(* IEC 61131-3 sources: volt/packages/volt-lsp-iec/test-corpus/lenze-mid/Device/Plc Logic/Application/Library Manager/CAA MemBlockMan, 94 files *)

(* ---- BCP.dut ---- *)
TYPE BCP :
STRUCT
	PPOOL : POINTER TO PCB;
END_STRUCT
END_TYPE

(* ---- ERROR.dut ---- *)
TYPE ERROR :
(
	NO_ERROR := 0,
	FIRST_ERROR := 30100,
	UNKNOWN_EVENT := 30102,
	NOMORE_MEMORY := 30103,
	WRONG_PRIO := 30104,
	EMPTY_LIST := 30105,
	NO_EXIST_PRIO := 30106,
	PRIO_EXIST := 30107,
	PRIOS_EXCEED := 30108,
	ALIGNMENT_ERROR := 30109,
	BLOCKSIZE_TO_SMALL := 30110,
	EMPTY_POOL := 30111,
	EMPTY_EXCHANGE := 30112,
	TIMEOUT := 30113,
	WRONG_TIMEOUT := 30114,
	REF_OVERFLOW := 30115,
	WRONG_KEY := 30116,
	HANDLE_INVALID := 30117,
	REF_NOT_ZERO := 30118,
	WRONG_NUM_OF_MSG := 30119,
	BUFFER_TO_BIG := 30120,
	WRONG_OP := 30121,
	GEN_ERROR := 30149,
	FIRST_MF := 30150,
	LAST_ERROR := 30199
);
END_TYPE

(* ---- PCB.dut ---- *)
TYPE PCB :
STRUCT
	XWDUMMYA : __XWORD;
	SZBLOCK : CAA.SIZE;
	XWDUMMYB : __XWORD;
	XWDUMMYC : __XWORD;
	CTBLKLEFT : CAA.COUNT;
	CTBLKCAP : CAA.COUNT;
END_STRUCT
END_TYPE

(* ---- RSHANDLING.gvl ---- *)
VAR_GLOBAL
	G_XCHGCLASS : XChgClass;
	G_FLATCLASS : FlatClass;
	G_MSGCLASS : MsgClass;
	G_REFCLASS : MsgClass;
	G_POOLCLASS : PoolClass;
	G_BLKCLASS : BlkClass;
	G_RLSTCLASS : RLstClass;
END_VAR

(* ---- VERSIONCONSTANTS.gvl ---- *)
VAR_GLOBAL
	GC_BYVERSION : BYTE := 1;
	GC_VERSION_1 : BYTE := 0;
END_VAR

(* ---- _BLOCKGETDATA.pou ---- *)
FUNCTION _BLOCKGETDATA : CAA.PVOID
VAR_INPUT
	HBLOCK : CAA.HANDLE;
	PEERROR : POINTER TO ERROR;
END_VAR
END_FUNCTION

(* ---- _BLOCKGETPOOL.pou ---- *)
FUNCTION _BLOCKGETPOOL : CAA.HANDLE
VAR_INPUT
	HBLOCK : CAA.HANDLE;
	PEERROR : POINTER TO ERROR;
END_VAR
END_FUNCTION

(* ---- _FLATCREATEH.pou ---- *)
FUNCTION _FLATCREATEH : CAA.HANDLE
VAR_INPUT
	IDMINKEY : CAA.IDENT;
	IDMAXKEY : CAA.IDENT;
	CTNUMKEYS : CAA.COUNT;
	EENABLE : CB.EVENT;
	EDISABLE : CB.EVENT;
	EUPDATE : CB.EVENT;
	EREAD : CB.EVENT;
	PEERROR : POINTER TO ERROR;
END_VAR
END_FUNCTION

(* ---- _FLATCREATEP.pou ---- *)
FUNCTION _FLATCREATEP : CAA.HANDLE
VAR_INPUT
	IDMINKEY : CAA.IDENT;
	IDMAXKEY : CAA.IDENT;
	CTNUMKEY : CAA.COUNT;
	SZMEMSIZE : CAA.SIZE;
	PMEMORY : CAA.PVOID;
	EENABLE : CB.EVENT;
	EDISABLE : CB.EVENT;
	EUPDATE : CB.EVENT;
	EREAD : CB.EVENT;
	PEERROR : POINTER TO ERROR;
END_VAR
END_FUNCTION

(* ---- _FLATDELETE.pou ---- *)
FUNCTION _FLATDELETE : ERROR
VAR_INPUT
	HFLAT : CAA.HANDLE;
END_VAR
END_FUNCTION

(* ---- _FLATDISABLE.pou ---- *)
FUNCTION _FLATDISABLE : CAA.HANDLE
VAR_INPUT
	HFLAT : CAA.HANDLE;
	IDKEY : CAA.IDENT;
	PEERROR : POINTER TO ERROR;
END_VAR
END_FUNCTION

(* ---- _FLATENABLE.pou ---- *)
FUNCTION _FLATENABLE : ERROR
VAR_INPUT
	HFLAT : CAA.HANDLE;
	IDKEY : CAA.IDENT;
END_VAR
END_FUNCTION

(* ---- _FLATGETSIZE.pou ---- *)
FUNCTION _FLATGETSIZE : CAA.SIZE
VAR_INPUT
	CTNUMKEYS : CAA.COUNT;
END_VAR
END_FUNCTION

(* ---- _FLATREAD.pou ---- *)
FUNCTION _FLATREAD : CAA.HANDLE
VAR_INPUT
	HFLAT : CAA.HANDLE;
	IDKEY : CAA.IDENT;
	PEERROR : POINTER TO ERROR;
END_VAR
END_FUNCTION

(* ---- _FLATTEST.pou ---- *)
FUNCTION _FLATTEST : BOOL
VAR_INPUT
	HFLAT : CAA.HANDLE;
	IDKEY : CAA.IDENT;
	PEERROR : POINTER TO ERROR;
END_VAR
END_FUNCTION

(* ---- _FLATUPDATE.pou ---- *)
FUNCTION _FLATUPDATE : CAA.HANDLE
VAR_INPUT
	HFLAT : CAA.HANDLE;
	IDKEY : CAA.IDENT;
	HMSG : CAA.HANDLE;
	PEERROR : POINTER TO ERROR;
END_VAR
END_FUNCTION

(* ---- _MSGADDREF.pou ---- *)
FUNCTION _MSGADDREF : ERROR
VAR_INPUT
	HMSG : CAA.HANDLE;
END_VAR
END_FUNCTION

(* ---- _MSGCLONE.pou ---- *)
FUNCTION _MSGCLONE : CAA.HANDLE
VAR_INPUT
	HMSG : CAA.HANDLE;
	PEERROR : POINTER TO ERROR;
END_VAR
END_FUNCTION

(* ---- _MSGGETDATA.pou ---- *)
FUNCTION _MSGGETDATA : CAA.PVOID
VAR_INPUT
	HMSG : CAA.HANDLE;
	PEERROR : POINTER TO ERROR;
END_VAR
END_FUNCTION

(* ---- _MSGRECEIVE.pou ---- *)
FUNCTION _MSGRECEIVE : CAA.HANDLE
VAR_INPUT
	HXCHG : CAA.HANDLE;
	PCTMSGLEFT : POINTER TO CAA.COUNT;
	PEERROR : POINTER TO ERROR;
END_VAR
END_FUNCTION

(* ---- _MSGRELEASE.pou ---- *)
FUNCTION _MSGRELEASE : ERROR
VAR_INPUT
	HMSG : CAA.HANDLE;
END_VAR
END_FUNCTION

(* ---- _MSGRELEASEEX.pou ---- *)
FUNCTION _MSGRELEASEEX : ERROR
VAR_INPUT
	HMSG : CAA.HANDLE;
	HXCHG : CAA.HANDLE;
END_VAR
END_FUNCTION

(* ---- _MSGSEND.pou ---- *)
FUNCTION _MSGSEND : ERROR
VAR_INPUT
	HMSG : CAA.HANDLE;
	USIPRIO : USINT;
	HXCHG : CAA.HANDLE;
END_VAR
END_FUNCTION

(* ---- _POOLCREATEH.pou ---- *)
FUNCTION _POOLCREATEH : CAA.HANDLE
VAR_INPUT
	CTNUMBLOCKS : CAA.COUNT;
	SZBLOCKSIZE : CAA.SIZE;
	EEMPTY : CB.EVENT;
	PEERROR : POINTER TO ERROR;
END_VAR
END_FUNCTION

(* ---- _POOLCREATEP.pou ---- *)
FUNCTION _POOLCREATEP : CAA.HANDLE
VAR_INPUT
	SZBLOCKSIZE : CAA.SIZE;
	SZMEMSIZE : CAA.SIZE;
	PMEMORY : CAA.PVOID;
	EEMPTY : CB.EVENT;
	PEERROR : POINTER TO ERROR;
END_VAR
END_FUNCTION

(* ---- _POOLDELETE.pou ---- *)
FUNCTION _POOLDELETE : ERROR
VAR_INPUT
	HPOOL : CAA.HANDLE;
END_VAR
END_FUNCTION

(* ---- _POOLEXTENDH.pou ---- *)
FUNCTION _POOLEXTENDH : ERROR
VAR_INPUT
	HPOOL : CAA.HANDLE;
	CTNUMBLOCKS : CAA.COUNT;
END_VAR
END_FUNCTION

(* ---- _POOLGETBLOCK.pou ---- *)
FUNCTION _POOLGETBLOCK : CAA.HANDLE
VAR_INPUT
	HPOOL : CAA.HANDLE;
	PEERROR : POINTER TO ERROR;
END_VAR
END_FUNCTION

(* ---- _POOLGETBLOCKSIZE.pou ---- *)
FUNCTION _POOLGETBLOCKSIZE : CAA.SIZE
VAR_INPUT
	HPOOL : CAA.HANDLE;
	PEERROR : POINTER TO ERROR;
END_VAR
END_FUNCTION

(* ---- _POOLGETCURCAPACITY.pou ---- *)
FUNCTION _POOLGETCURCAPACITY : CAA.COUNT
VAR_INPUT
	HPOOL : CAA.HANDLE;
	PEERROR : POINTER TO ERROR;
END_VAR
END_FUNCTION

(* ---- _POOLGETNUMBLOCKSLEFT.pou ---- *)
FUNCTION _POOLGETNUMBLOCKSLEFT : CAA.COUNT
VAR_INPUT
	HPOOL : CAA.HANDLE;
	PEERROR : POINTER TO ERROR;
END_VAR
END_FUNCTION

(* ---- _POOLGETSIZE.pou ---- *)
FUNCTION _POOLGETSIZE : CAA.SIZE
VAR_INPUT
	CTNUMBLOCK : CAA.COUNT;
	SZBLOCKSIZE : CAA.SIZE;
END_VAR
END_FUNCTION

(* ---- _POOLPUTBLOCK.pou ---- *)
FUNCTION _POOLPUTBLOCK : ERROR
VAR_INPUT
	HBLOCK : CAA.HANDLE;
END_VAR
END_FUNCTION

(* ---- _RLSTADDPRIO.pou ---- *)
FUNCTION _RLSTADDPRIO : ERROR
VAR_INPUT
	HRLST : CAA.HANDLE;
	USIPRIO : USINT;
END_VAR
END_FUNCTION

(* ---- _RLSTCHECKPRIO.pou ---- *)
FUNCTION _RLSTCHECKPRIO : BOOL
VAR_INPUT
	HRLST : CAA.HANDLE;
	USIPRIO : USINT;
	PEERROR : POINTER TO ERROR;
END_VAR
END_FUNCTION

(* ---- _RLSTCREATEH.pou ---- *)
FUNCTION _RLSTCREATEH : CAA.HANDLE
VAR_INPUT
	PEERROR : POINTER TO ERROR;
END_VAR
END_FUNCTION

(* ---- _RLSTCREATEP.pou ---- *)
FUNCTION _RLSTCREATEP : CAA.HANDLE
VAR_INPUT
	SZMEMORY : CAA.SIZE;
	PMEMORY : CAA.PVOID;
	PEERROR : POINTER TO ERROR;
END_VAR
END_FUNCTION

(* ---- _RLSTDELETE.pou ---- *)
FUNCTION _RLSTDELETE : ERROR
VAR_INPUT
	HRLST : CAA.HANDLE;
END_VAR
END_FUNCTION

(* ---- _RLSTGETHIGHESTPRIO.pou ---- *)
FUNCTION _RLSTGETHIGHESTPRIO : USINT
VAR_INPUT
	HRLST : CAA.HANDLE;
	PEERROR : POINTER TO ERROR;
END_VAR
END_FUNCTION

(* ---- _RLSTGETSIZE.pou ---- *)
FUNCTION _RLSTGETSIZE : CAA.SIZE
VAR_INPUT
	XDUMMY : BOOL;
END_VAR
END_FUNCTION

(* ---- _RLSTREMOVEPRIO.pou ---- *)
FUNCTION _RLSTREMOVEPRIO : ERROR
VAR_INPUT
	HRLST : CAA.HANDLE;
	USIPRIO : USINT;
END_VAR
END_FUNCTION

(* ---- _XCHGCREATEH.pou ---- *)
FUNCTION _XCHGCREATEH : CAA.HANDLE
VAR_INPUT
	CTNUMMSG : CAA.COUNT;
	SZBLOCKSIZE : CAA.SIZE;
	CTNUMPRIOS : CAA.COUNT;
	ESENDMSG : CB.EVENT;
	ERECEIVEMSG : CB.EVENT;
	EXCHGEMPTY : CB.EVENT;
	PEERROR : POINTER TO ERROR;
END_VAR
END_FUNCTION

(* ---- _XCHGCREATEP.pou ---- *)
FUNCTION _XCHGCREATEP : CAA.HANDLE
VAR_INPUT
	SZBLOCKSIZE : CAA.SIZE;
	CTNUMPRIOS : CAA.COUNT;
	SZMEMSIZE : CAA.SIZE;
	PMEMORY : CAA.PVOID;
	ESENDMSG : CB.EVENT;
	ERECEIVEMSG : CB.EVENT;
	EXCHGEMPTY : CB.EVENT;
	PEERROR : POINTER TO ERROR;
END_VAR
END_FUNCTION

(* ---- _XCHGDELETE.pou ---- *)
FUNCTION _XCHGDELETE : ERROR
VAR_INPUT
	HXCHG : CAA.HANDLE;
END_VAR
END_FUNCTION

(* ---- _XCHGEXTENDH.pou ---- *)
FUNCTION _XCHGEXTENDH : ERROR
VAR_INPUT
	HXCHG : CAA.HANDLE;
	CTNUMMSG : CAA.COUNT;
END_VAR
END_FUNCTION

(* ---- _XCHGGETSIZE.pou ---- *)
FUNCTION _XCHGGETSIZE : CAA.SIZE
VAR_INPUT
	CTNUMMSG : CAA.COUNT;
	SZBLOCKSIZE : CAA.SIZE;
	CTNUMPRIOS : CAA.COUNT;
END_VAR
END_FUNCTION

(* ---- _XCHGISEMPTY.pou ---- *)
FUNCTION _XCHGISEMPTY : BOOL
VAR_INPUT
	HXCHG : CAA.HANDLE;
	PEERROR : POINTER TO ERROR;
END_VAR
END_FUNCTION

(* ---- _XCHGMSGLEFT.pou ---- *)
FUNCTION _XCHGMSGLEFT : CAA.COUNT
VAR_INPUT
	HXCHG : CAA.HANDLE;
	PEERROR : POINTER TO ERROR;
END_VAR
END_FUNCTION

(* ---- BLOCKGETDATA.pou ---- *)
FUNCTION BLOCKGETDATA : CAA.PVOID
VAR_INPUT
	HBLOCK : CAA.HANDLE;
	PEERROR : POINTER TO ERROR;
END_VAR
END_FUNCTION

(* ---- FLATCREATEH.pou ---- *)
FUNCTION FLATCREATEH : CAA.HANDLE
VAR_INPUT
	IDMINKEY : CAA.IDENT;
	IDMAXKEY : CAA.IDENT;
	CTNUMKEYS : CAA.COUNT;
	EENABLE : CB.EVENT;
	EDISABLE : CB.EVENT;
	EUPDATE : CB.EVENT;
	EREAD : CB.EVENT;
	PEERROR : POINTER TO ERROR;
END_VAR
END_FUNCTION

(* ---- FLATCREATEP.pou ---- *)
FUNCTION FLATCREATEP : CAA.HANDLE
VAR_INPUT
	IDMINKEY : CAA.IDENT;
	IDMAXKEY : CAA.IDENT;
	CTNUMKEY : CAA.COUNT;
	SZMEMSIZE : CAA.SIZE;
	PMEMORY : CAA.PVOID;
	EENABLE : CB.EVENT;
	EDISABLE : CB.EVENT;
	EUPDATE : CB.EVENT;
	EREAD : CB.EVENT;
	PEERROR : POINTER TO ERROR;
END_VAR
END_FUNCTION

(* ---- FLATDELETE.pou ---- *)
FUNCTION FLATDELETE : ERROR
VAR_INPUT
	HFLAT : CAA.HANDLE;
END_VAR
END_FUNCTION

(* ---- FLATDISABLE.pou ---- *)
FUNCTION FLATDISABLE : CAA.HANDLE
VAR_INPUT
	HFLAT : CAA.HANDLE;
	IDKEY : CAA.IDENT;
	PEERROR : POINTER TO ERROR;
END_VAR
END_FUNCTION

(* ---- FLATENABLE.pou ---- *)
FUNCTION FLATENABLE : ERROR
VAR_INPUT
	HFLAT : CAA.HANDLE;
	IDKEY : CAA.IDENT;
END_VAR
END_FUNCTION

(* ---- FLATGETSIZE.pou ---- *)
FUNCTION FLATGETSIZE : CAA.SIZE
VAR_INPUT
	CTNUMKEYS : CAA.COUNT;
END_VAR
END_FUNCTION

(* ---- FLATREAD.pou ---- *)
FUNCTION FLATREAD : CAA.HANDLE
VAR_INPUT
	HFLAT : CAA.HANDLE;
	IDKEY : CAA.IDENT;
	PEERROR : POINTER TO ERROR;
END_VAR
END_FUNCTION

(* ---- FLATTEST.pou ---- *)
FUNCTION FLATTEST : BOOL
VAR_INPUT
	HFLAT : CAA.HANDLE;
	IDKEY : CAA.IDENT;
	PEERROR : POINTER TO ERROR;
END_VAR
END_FUNCTION

(* ---- FLATUPDATE.pou ---- *)
FUNCTION FLATUPDATE : CAA.HANDLE
VAR_INPUT
	HFLAT : CAA.HANDLE;
	IDKEY : CAA.IDENT;
	HMSG : CAA.HANDLE;
	PEERROR : POINTER TO ERROR;
END_VAR
END_FUNCTION

(* ---- GETSUPPLIERVERSION.pou ---- *)
FUNCTION GETSUPPLIERVERSION : WORD
VAR_INPUT
	XDUMMY : BOOL;
END_VAR
END_FUNCTION

(* ---- MSGADDREF.pou ---- *)
FUNCTION MSGADDREF : ERROR
VAR_INPUT
	HMSG : CAA.HANDLE;
END_VAR
END_FUNCTION

(* ---- MSGCLONE.pou ---- *)
FUNCTION MSGCLONE : CAA.HANDLE
VAR_INPUT
	HMSG : CAA.HANDLE;
	PEERROR : POINTER TO ERROR;
END_VAR
END_FUNCTION

(* ---- MSGGETDATA.pou ---- *)
FUNCTION MSGGETDATA : CAA.PVOID
VAR_INPUT
	HMSG : CAA.HANDLE;
	PEERROR : POINTER TO ERROR;
END_VAR
END_FUNCTION

(* ---- MSGRECEIVE.pou ---- *)
FUNCTION MSGRECEIVE : CAA.HANDLE
VAR_INPUT
	HXCHG : CAA.HANDLE;
	PCTMSGLEFT : POINTER TO CAA.COUNT;
	PEERROR : POINTER TO ERROR;
END_VAR
END_FUNCTION

(* ---- MSGRELEASE.pou ---- *)
FUNCTION MSGRELEASE : ERROR
VAR_INPUT
	HMSG : CAA.HANDLE;
END_VAR
END_FUNCTION

(* ---- MSGRELEASEEX.pou ---- *)
FUNCTION MSGRELEASEEX : ERROR
VAR_INPUT
	HMSG : CAA.HANDLE;
	HXCHG : CAA.HANDLE;
END_VAR
END_FUNCTION

(* ---- MSGSEND.pou ---- *)
FUNCTION MSGSEND : ERROR
VAR_INPUT
	HMSG : CAA.HANDLE;
	USIPRIO : USINT;
	HXCHG : CAA.HANDLE;
END_VAR
END_FUNCTION

(* ---- POOLCREATEH.pou ---- *)
FUNCTION POOLCREATEH : CAA.HANDLE
VAR_INPUT
	CTNUMBLOCKS : CAA.COUNT;
	SZBLOCKSIZE : CAA.SIZE;
	EEMPTY : CB.EVENT;
	PEERROR : POINTER TO ERROR;
END_VAR
END_FUNCTION

(* ---- POOLCREATEP.pou ---- *)
FUNCTION POOLCREATEP : CAA.HANDLE
VAR_INPUT
	SZBLOCKSIZE : CAA.SIZE;
	SZMEMSIZE : CAA.SIZE;
	PMEMORY : CAA.PVOID;
	EEMPTY : CB.EVENT;
	PEERROR : POINTER TO ERROR;
END_VAR
END_FUNCTION

(* ---- POOLDELETE.pou ---- *)
FUNCTION POOLDELETE : ERROR
VAR_INPUT
	HPOOL : CAA.HANDLE;
END_VAR
END_FUNCTION

(* ---- POOLEXTENDH.pou ---- *)
FUNCTION POOLEXTENDH : ERROR
VAR_INPUT
	HPOOL : CAA.HANDLE;
	CTNUMBLOCKS : CAA.COUNT;
END_VAR
END_FUNCTION

(* ---- POOLGETBLOCK.pou ---- *)
FUNCTION POOLGETBLOCK : CAA.HANDLE
VAR_INPUT
	HPOOL : CAA.HANDLE;
	PEERROR : POINTER TO ERROR;
END_VAR
END_FUNCTION

(* ---- POOLGETSIZE.pou ---- *)
FUNCTION POOLGETSIZE : CAA.SIZE
VAR_INPUT
	CTNUMBLOCK : CAA.COUNT;
	SZBLOCKSIZE : CAA.SIZE;
END_VAR
END_FUNCTION

(* ---- POOLPUTBLOCK.pou ---- *)
FUNCTION POOLPUTBLOCK : ERROR
VAR_INPUT
	HBLOCK : CAA.HANDLE;
END_VAR
END_FUNCTION

(* ---- RLSTADDPRIO.pou ---- *)
FUNCTION RLSTADDPRIO : ERROR
VAR_INPUT
	HRLST : CAA.HANDLE;
	USIPRIO : USINT;
END_VAR
END_FUNCTION

(* ---- RLSTCHECKPRIO.pou ---- *)
FUNCTION RLSTCHECKPRIO : BOOL
VAR_INPUT
	HRLST : CAA.HANDLE;
	USIPRIO : USINT;
	PEERROR : POINTER TO ERROR;
END_VAR
END_FUNCTION

(* ---- RLSTCREATEH.pou ---- *)
FUNCTION RLSTCREATEH : CAA.HANDLE
VAR_INPUT
	PEERROR : POINTER TO ERROR;
END_VAR
END_FUNCTION

(* ---- RLSTCREATEP.pou ---- *)
FUNCTION RLSTCREATEP : CAA.HANDLE
VAR_INPUT
	SZMEMORY : CAA.SIZE;
	PMEMORY : CAA.PVOID;
	PEERROR : POINTER TO ERROR;
END_VAR
END_FUNCTION

(* ---- RLSTDELETE.pou ---- *)
FUNCTION RLSTDELETE : ERROR
VAR_INPUT
	HRLST : CAA.HANDLE;
END_VAR
END_FUNCTION

(* ---- RLSTGETHIGHESTPRIO.pou ---- *)
FUNCTION RLSTGETHIGHESTPRIO : USINT
VAR_INPUT
	HRLST : CAA.HANDLE;
	PEERROR : POINTER TO ERROR;
END_VAR
END_FUNCTION

(* ---- RLSTGETSIZE.pou ---- *)
FUNCTION RLSTGETSIZE : CAA.SIZE
VAR_INPUT
	XDUMMY : BOOL;
END_VAR
END_FUNCTION

(* ---- RLSTREMOVEPRIO.pou ---- *)
FUNCTION RLSTREMOVEPRIO : ERROR
VAR_INPUT
	HRLST : CAA.HANDLE;
	USIPRIO : USINT;
END_VAR
END_FUNCTION

(* ---- XCHGCREATEH.pou ---- *)
FUNCTION XCHGCREATEH : CAA.HANDLE
VAR_INPUT
	CTNUMMSG : CAA.COUNT;
	SZBLOCKSIZE : CAA.SIZE;
	CTNUMPRIOS : CAA.COUNT;
	ESENDMSG : CB.EVENT;
	ERECEIVEMSG : CB.EVENT;
	EXCHGEMPTY : CB.EVENT;
	PEERROR : POINTER TO ERROR;
END_VAR
END_FUNCTION

(* ---- XCHGCREATEP.pou ---- *)
FUNCTION XCHGCREATEP : CAA.HANDLE
VAR_INPUT
	SZBLOCKSIZE : CAA.SIZE;
	CTNUMPRIOS : CAA.COUNT;
	SZMEMSIZE : CAA.SIZE;
	PMEMORY : CAA.PVOID;
	ESENDMSG : CB.EVENT;
	ERECEIVEMSG : CB.EVENT;
	EXCHGEMPTY : CB.EVENT;
	PEERROR : POINTER TO ERROR;
END_VAR
END_FUNCTION

(* ---- XCHGDELETE.pou ---- *)
FUNCTION XCHGDELETE : ERROR
VAR_INPUT
	HXCHG : CAA.HANDLE;
END_VAR
END_FUNCTION

(* ---- XCHGEXTENDH.pou ---- *)
FUNCTION XCHGEXTENDH : ERROR
VAR_INPUT
	HXCHG : CAA.HANDLE;
	CTNUMMSG : CAA.COUNT;
END_VAR
END_FUNCTION

(* ---- XCHGGETSIZE.pou ---- *)
FUNCTION XCHGGETSIZE : CAA.SIZE
VAR_INPUT
	CTNUMMSG : CAA.COUNT;
	SZBLOCKSIZE : CAA.SIZE;
	CTNUMPRIOS : CAA.COUNT;
END_VAR
END_FUNCTION

(* ---- XCHGISEMPTY.pou ---- *)
FUNCTION XCHGISEMPTY : BOOL
VAR_INPUT
	HXCHG : CAA.HANDLE;
	PEERROR : POINTER TO ERROR;
END_VAR
END_FUNCTION

(* ---- XCHGMSGLEFT.pou ---- *)
FUNCTION XCHGMSGLEFT : CAA.COUNT
VAR_INPUT
	HXCHG : CAA.HANDLE;
	PEERROR : POINTER TO ERROR;
END_VAR
END_FUNCTION

(* ---- BLKCLASS.pou ---- *)
FUNCTION_BLOCK BLKCLASS EXTENDS RSMClass
END_FUNCTION_BLOCK

METHOD CLOSE : RSM.ERROR
VAR_INPUT
	HHANDLE : CAA.HANDLE;
END_VAR
END_METHOD

(* ---- FLATCLASS.pou ---- *)
FUNCTION_BLOCK FLATCLASS EXTENDS RSMClass
END_FUNCTION_BLOCK

METHOD CLOSE : RSM.ERROR
VAR_INPUT
	HHANDLE : CAA.HANDLE;
END_VAR
END_METHOD

(* ---- MSGCLASS.pou ---- *)
FUNCTION_BLOCK MSGCLASS EXTENDS RSMClass
END_FUNCTION_BLOCK

METHOD CLOSE : RSM.ERROR
VAR_INPUT
	HHANDLE : CAA.HANDLE;
END_VAR
END_METHOD

(* ---- POOLCLASS.pou ---- *)
FUNCTION_BLOCK POOLCLASS EXTENDS RSMClass
END_FUNCTION_BLOCK

METHOD CLOSE : RSM.ERROR
VAR_INPUT
	HHANDLE : CAA.HANDLE;
END_VAR
END_METHOD

(* ---- RLSTCLASS.pou ---- *)
FUNCTION_BLOCK RLSTCLASS EXTENDS RSMClass
END_FUNCTION_BLOCK

METHOD CLOSE : RSM.ERROR
VAR_INPUT
	HHANDLE : CAA.HANDLE;
END_VAR
END_METHOD

(* ---- XCHGCLASS.pou ---- *)
FUNCTION_BLOCK XCHGCLASS EXTENDS RSMClass
END_FUNCTION_BLOCK

METHOD CLOSE : RSM.ERROR
VAR_INPUT
	HHANDLE : CAA.HANDLE;
END_VAR
END_METHOD
